TYPE ST_Val :
STRUCT
	fValue		: REAL;
	bValid		: BOOL;		// FALSE면 fValue를 쓰지 않는다
END_STRUCT
END_TYPE

(* stored: Version 1.1.0.1, ProductVersion 3.1.4024.15
   DUT ST_Val: Id {aa4e7fde-9b80-4f72-854c-7a4f3cbd81e4} *)
